SUBAPPLICATION Boot_Zaehler_OPC (* STG1: meldet READY=TRUE und nimmt Boot-Meldungen der Stationen per Methode entgegen (Argument = STG-Nummer) *)
  (* Standard: 61499-2; Description: Copyright (c) 2026 Meisterschulen am Ostbahnhof This program and the accompanying materials are made available under the terms of the Eclipse Public License 2.0 which is available at https://www.eclipse.org/legal/epl-2.0/ SPDX-License-Identifier: EPL-2.0 *)
  (* Version 1.1, 2026-11-25, Franz Höpfinger, Meisterschulen am Ostbahnhof, IND nur bei QO=TRUE an RSP und Verteiler (E_PERMIT). Ein gescheitertes RSP meldet IND mit QO=FALSE, direkt IND->RSP ergab eine Endlosschleife (Zaehler STG4 lief hoch, STG3 rot). *)
  (* Version 1.0, 2026-10-29, Franz Höpfinger, Meisterschulen am Ostbahnhof, Neu (Franz: STG1 verwaltet alle Boot-Zaehler, ohne INI). READY wird bei INIT einmal TRUE publiziert, die Stationen rufen bei steigender Flanke die Methode mit ihrer Nummer auf (Boot_Melden_OPC). E_DEMUX_6 verteilt K=2..5 auf BOOT_STG2..5. *)
  PACKAGE MyLib::sys;
  (* Documentation:
  Boot-Zähler auf STG1
   STG1 veröffentlicht nach dem Start einmal READY = TRUE. STG2–5 abonnieren diesen Wert (Boot_Melden_OPC). Sobald eine Station TRUE sieht (steigende Flanke nach ihrem eigenen Start), ruft sie die Methode BOOT_MELDUNG mit ihrer STG-Nummer auf. Ein reiner Verbindungsabbruch löst keine Flanke aus, nur ein Neustart der Station.
   Gezählt wird in Station_Alive_VT_OPC (Eingang BOOT), nur im RAM, ohne INI.
   IND geht nur bei QO = TRUE an RSP und den Verteiler (E_PERMIT). Findet FORTE zu einem RSP keinen offenen Aufruf (z. B. nach dem 4-s-Timeout), meldet der SERVER IND mit QO = FALSE und altem RD_1. Direkt IND→RSP verdrahtet ergibt das eine Endlosschleife.
  *)
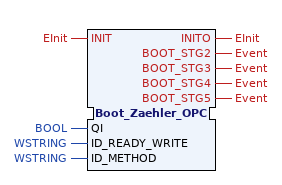
  EVENT_INPUT
    INIT : EInit; (* Initialization Request *)
  END_EVENT
  EVENT_OUTPUT
    INITO : EInit; (* Initialization Confirm *)
    BOOT_STG2; (* STG2 ist gestartet *)
    BOOT_STG3; (* STG3 ist gestartet *)
    BOOT_STG4; (* STG4 ist gestartet *)
    BOOT_STG5; (* STG5 ist gestartet *)
  END_EVENT
  VAR_INPUT
    QI : BOOL := TRUE; (* Quality Input - TRUE to enable service *)
    ID_READY_WRITE : WSTRING; (* Lokaler Knoten READY (BOOL) *)
    ID_METHOD : WSTRING; (* Lokale Methode BOOT_MELDUNG (1 UINT-Argument) *)
  END_VAR
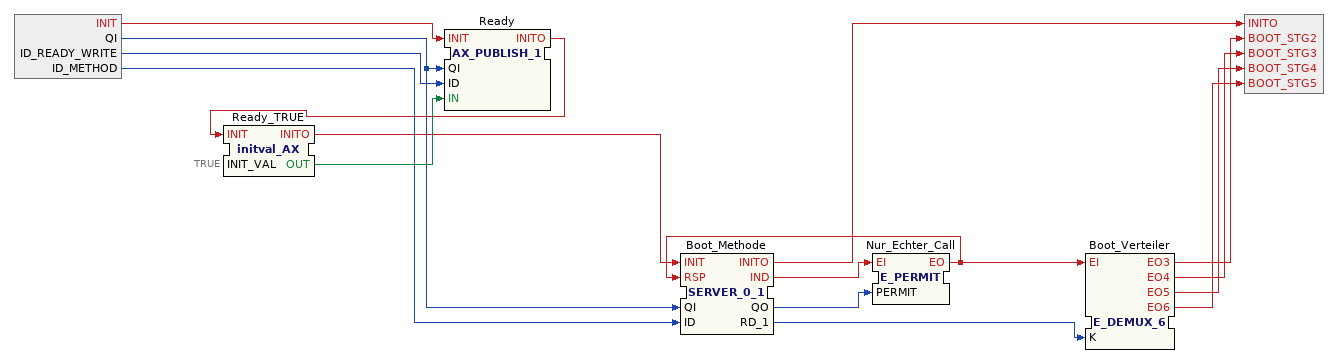
  FBS
    Ready : adapter::net::AX_PUBLISH_1;
    Ready_TRUE : adapter::types::unidirectional::AX::initval::initval_AX(INIT_VAL := TRUE);
    Boot_Methode : iec61499::net::SERVER_0_1; (* IND->RSP nur bei QO *)
    Nur_Echter_Call : iec61499::events::E_PERMIT; (* nur echter Call (QO=TRUE) *)
    Boot_Verteiler : iec61499::events::E_DEMUX_6; (* K = STG-Nummer *)
  END_FBS
  EVENT_CONNECTIONS
    INIT TO Ready.INIT;
    Ready.INITO TO Ready_TRUE.INIT;
    Ready_TRUE.INITO TO Boot_Methode.INIT;
    Boot_Methode.INITO TO INITO;
    Boot_Methode.IND TO Nur_Echter_Call.EI;
    Nur_Echter_Call.EO TO Boot_Methode.RSP;
    Nur_Echter_Call.EO TO Boot_Verteiler.EI;
    Boot_Verteiler.EO3 TO BOOT_STG2;
    Boot_Verteiler.EO4 TO BOOT_STG3;
    Boot_Verteiler.EO5 TO BOOT_STG4;
    Boot_Verteiler.EO6 TO BOOT_STG5;
  END_CONNECTIONS
  DATA_CONNECTIONS
    QI TO Ready.QI;
    ID_READY_WRITE TO Ready.ID;
    QI TO Boot_Methode.QI;
    ID_METHOD TO Boot_Methode.ID;
    Boot_Methode.QO TO Nur_Echter_Call.PERMIT;
    Boot_Methode.RD_1 TO Boot_Verteiler.K;
  END_CONNECTIONS
  ADAPTER_CONNECTIONS
    Ready_TRUE.OUT TO Ready.IN;
  END_CONNECTIONS
END_SUBAPPLICATION
